// TIA Portal V21 export
// export: Created 2026-11-11T00:47:19.431695Z, ExportSetting WithDefaults, DisplayName Totally Integrated Automation Portal, DisplayVersion V21 Update 3, DisplayName STEP 7 Professional, DisplayVersion V21 Update 3, DisplayName STEP 7 Safety, DisplayVersion V21, DisplayName Tech WebApplication, DisplayVersion V21, DisplayName WinCC Basic/Comfort/Advanced, DisplayVersion V21 Update 3, DisplayName WinCC Unified, DisplayVersion V21 Update 3
FUNCTION_BLOCK "FB_Fbd_ex056"   // FB94, FBD
{ S7_Optimized_Access := 'TRUE' }
VERSION : 0.1
// stored: AutoNumber true, IsIECCheckEnabled false, IsRetainMemResEnabled false, MemoryReserve 100, SetENOAutomatically false, UDAEnableTagReadback false
   VAR_INPUT
      v_req : Bool;
      v_mode : USInt;
      v_laddr : HW_DEVICE;
   END_VAR
   VAR_OUTPUT
      v_ret_val : Int;
      v_busy : Bool;
   END_VAR
BEGIN

REGION Network 1: D_ACT_DP - Activate/deactivate DP slaves
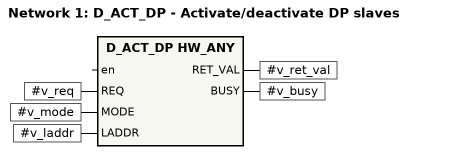
   #v_ret_val := D_ACT_DP(REQ := #v_req, MODE := #v_mode, LADDR := #v_laddr, BUSY => #v_busy);
END_REGION
END_FUNCTION_BLOCK
